Fanuc KAREL source: kc00043.KL

-- PROVISIONAL review KL for V1013-1; original PC SHA256 638eb59bea7ebc35e1e971eb06c540d1f8a1b1c21ab1211c3a013a293e8579f5
-- Incomplete behavior may be omitted. Consult companion uncertainty JSON. Do not deploy.
PROGRAM KC00043
%NOLOCKGROUP
BEGIN
  -- UNRESOLVED_PC offsets 5-35; opcodes 27,22,22,27,9D,31,7E,4A
  -- UNRESOLVED_PC offsets 40-44; opcodes 7F
END KC00043
